// TIA Portal V20 export
DATA_BLOCK "DB_Stoermeldungen"   // DB512
TITLE = Schnittstelle OP_AG 1
{ S7_Optimized_Access := 'FALSE' }
AUTHOR : SD
FAMILY : KOMM
// stored: AutoNumber false
   VAR RETAIN
      Allgemeine { S7_SetPoint := 'True'} : "Störmeldung";
      Allgemeine_1 { S7_SetPoint := 'True'} : "Störmeldung";
      SM_Wartungszähler { S7_SetPoint := 'True'} : "Störmeldung";
      Störmeldungen_PN : "Störmeldung_PN";
   END_VAR
BEGIN
   Allgemeine.Störmeldung[0] := FALSE;
   Allgemeine.Störmeldung[1] := FALSE;   // SM1 Systemdruck nicht vorhanden ! Prüfen und Weiter mit ACK
   Allgemeine.Störmeldung[2] := FALSE;   // SM2 Anlagendruck nicht aufgebaut -939S1
   Allgemeine.Störmeldung[3] := FALSE;   // SM3 Algemein Richten Gesamtanlage erforderlich
   Allgemeine.Störmeldung[4] := FALSE;   // SM4 Richten Gesamtanlage nach Teil neu geladen
   Allgemeine.Störmeldung[5] := FALSE;   // SM5
   Allgemeine.Störmeldung[6] := FALSE;   // SM6
   Allgemeine.Störmeldung[7] := FALSE;   // SM7
   Allgemeine.Störmeldung[8] := FALSE;   // SM8
   Allgemeine.Störmeldung[9] := FALSE;   // SM9
   Allgemeine.Störmeldung[10] := FALSE;   // SM10
   Allgemeine.Störmeldung[11] := FALSE;   // SM11
   Allgemeine.Störmeldung[12] := FALSE;   // SM12
   Allgemeine.Störmeldung[13] := FALSE;   // SM13
   Allgemeine.Störmeldung[14] := FALSE;   // SM14
   Allgemeine.Störmeldung[15] := FALSE;   // SM15
   Allgemeine.Störmeldung[16] := FALSE;   // SM16
   Allgemeine.Störmeldung[17] := FALSE;   // SM17
   Allgemeine.Störmeldung[18] := FALSE;   // SM18
   Allgemeine.Störmeldung[19] := FALSE;   // SM19
   Allgemeine.Störmeldung[20] := FALSE;   // SM20
   Allgemeine.Störmeldung[21] := FALSE;   // SM21
   Allgemeine.Störmeldung[22] := FALSE;   // SM22
   Allgemeine.Störmeldung[23] := FALSE;   // SM23
   Allgemeine.Störmeldung[24] := FALSE;   // SM24
   Allgemeine.Störmeldung[25] := FALSE;   // SM25
   Allgemeine.Störmeldung[26] := FALSE;   // SM26
   Allgemeine.Störmeldung[27] := FALSE;   // SM27
   Allgemeine.Störmeldung[28] := FALSE;   // SM28
   Allgemeine.Störmeldung[29] := FALSE;   // SM29
   Allgemeine.Störmeldung[30] := FALSE;   // SM30
   Allgemeine.Störmeldung[31] := FALSE;   // SM31
   Allgemeine_1.Störmeldung[0] := FALSE;   // SM32 Schutztüre 1 nicht verriegelt
   Allgemeine_1.Störmeldung[1] := FALSE;   // SM33 Schutztüre 2 nicht verriegelt
   Allgemeine_1.Störmeldung[2] := FALSE;   // SM34 Schutztüre 3 nicht verriegelt
   Allgemeine_1.Störmeldung[3] := FALSE;   // SM35 Schutztüre 4 nicht verriegelt
   Allgemeine_1.Störmeldung[4] := FALSE;   // SM36 Schutztüre 5 nicht verriegelt
   Allgemeine_1.Störmeldung[5] := FALSE;   // SM37 Schutztüre 6 nicht verriegelt
   Allgemeine_1.Störmeldung[6] := FALSE;   // SM38 Schutztüre 7 nicht verriegelt
   Allgemeine_1.Störmeldung[7] := FALSE;   // SM39 Schutztüre 8 nicht verriegelt
   Allgemeine_1.Störmeldung[8] := FALSE;   // SM40 Schutztüre 9 nicht verriegelt
   Allgemeine_1.Störmeldung[9] := FALSE;   // SM41 Schutztüre 10 nicht verriegelt
   Allgemeine_1.Störmeldung[10] := FALSE;   // SM42 Schutztüre 11 nicht verriegelt
   Allgemeine_1.Störmeldung[11] := FALSE;   // SM43 Steuerspannung 24V nicht in Ordnung
   Allgemeine_1.Störmeldung[12] := FALSE;   // SM44 Not-Aus Taster Bedienpanel
   Allgemeine_1.Störmeldung[13] := FALSE;   // SM45 Not-Aus Taster extern
   Allgemeine_1.Störmeldung[14] := FALSE;   // SM46 Kontrolle Box 1 voll -> leeren -> Start
   Allgemeine_1.Störmeldung[15] := FALSE;   // SM47 Kontrolle Box 2 voll -> leeren -> Start
   Allgemeine_1.Störmeldung[16] := FALSE;   // SM48 Kontrolle Box 3 voll -> leeren -> Start
   Allgemeine_1.Störmeldung[17] := FALSE;   // SM49 NIO Box 1 voll -> leeren -> Start
   Allgemeine_1.Störmeldung[18] := FALSE;   // SM50 NIO Box 2 voll -> leeren -> Start
   Allgemeine_1.Störmeldung[19] := FALSE;   // SM51 IO Box voll -> leeren -> Start
   Allgemeine_1.Störmeldung[20] := FALSE;   // SM52 Teiledaten wurden nicht richtig übertragen
   Allgemeine_1.Störmeldung[21] := FALSE;   // SM53 IO Box in Einhausung voll -> leeren -> Start
   Allgemeine_1.Störmeldung[22] := FALSE;   // SM54
   Allgemeine_1.Störmeldung[23] := FALSE;   // SM55 Anlagendruck bei Not-Halt nicht abgebaut -939S2
   Allgemeine_1.Störmeldung[24] := FALSE;   // SM56 Überspannungsschutz nicht OK
   Allgemeine_1.Störmeldung[25] := FALSE;   // SM57
   Allgemeine_1.Störmeldung[26] := FALSE;   // SM58
   Allgemeine_1.Störmeldung[27] := FALSE;   // SM59
   Allgemeine_1.Störmeldung[28] := FALSE;   // SM60
   Allgemeine_1.Störmeldung[29] := FALSE;   // SM61
   Allgemeine_1.Störmeldung[30] := FALSE;   // SM62
   Allgemeine_1.Störmeldung[31] := FALSE;   // SM63
   SM_Wartungszähler.Störmeldung[0] := FALSE;   // SM576 Wartungszähler 1
   SM_Wartungszähler.Störmeldung[1] := FALSE;   // SM577 Wartungszähler 2
   SM_Wartungszähler.Störmeldung[2] := FALSE;   // SM578 Wartungszähler 3
   SM_Wartungszähler.Störmeldung[3] := FALSE;   // SM579 Wartungszähler 4
   SM_Wartungszähler.Störmeldung[4] := FALSE;   // SM580 Wartungszähler 5
   SM_Wartungszähler.Störmeldung[5] := FALSE;   // SM581 Wartungszähler 6
   SM_Wartungszähler.Störmeldung[6] := FALSE;   // SM582 Wartungszähler 7
   SM_Wartungszähler.Störmeldung[7] := FALSE;   // SM583
   SM_Wartungszähler.Störmeldung[8] := FALSE;   // SM584
   SM_Wartungszähler.Störmeldung[9] := FALSE;   // SM585
   SM_Wartungszähler.Störmeldung[10] := FALSE;   // SM586
   SM_Wartungszähler.Störmeldung[11] := FALSE;   // SM587
   SM_Wartungszähler.Störmeldung[12] := FALSE;   // SM588
   SM_Wartungszähler.Störmeldung[13] := FALSE;   // SM589
   SM_Wartungszähler.Störmeldung[14] := FALSE;   // SM590
   SM_Wartungszähler.Störmeldung[15] := FALSE;   // SM591
   SM_Wartungszähler.Störmeldung[16] := FALSE;   // SM592
   SM_Wartungszähler.Störmeldung[17] := FALSE;   // SM593
   SM_Wartungszähler.Störmeldung[18] := FALSE;   // SM594
   SM_Wartungszähler.Störmeldung[19] := FALSE;   // SM595
   SM_Wartungszähler.Störmeldung[20] := FALSE;   // SM596
   SM_Wartungszähler.Störmeldung[21] := FALSE;   // SM597
   SM_Wartungszähler.Störmeldung[22] := FALSE;   // SM598
   SM_Wartungszähler.Störmeldung[23] := FALSE;   // SM599
   SM_Wartungszähler.Störmeldung[24] := FALSE;   // SM600
   SM_Wartungszähler.Störmeldung[25] := FALSE;   // SM601
   SM_Wartungszähler.Störmeldung[26] := FALSE;   // SM602
   SM_Wartungszähler.Störmeldung[27] := FALSE;   // SM603
   SM_Wartungszähler.Störmeldung[28] := FALSE;   // SM604
   SM_Wartungszähler.Störmeldung[29] := FALSE;   // SM605
   SM_Wartungszähler.Störmeldung[30] := FALSE;   // SM606
   SM_Wartungszähler.Störmeldung[31] := FALSE;   // SM607
   Störmeldungen_PN.Störmeldung_PN[0] := FALSE;   // SM608 Sammelstörung Profinet
   Störmeldungen_PN.Störmeldung_PN[1] := FALSE;   // SM609 Ausfall/Störung +HS1-101A1 Pluto Gateway Profinet
   Störmeldungen_PN.Störmeldung_PN[2] := FALSE;   // SM610 Ausfall/Störung +HS1-41T1 Pos 3.0 Drehteller
   Störmeldungen_PN.Störmeldung_PN[3] := FALSE;   // SM611 Ausfall/Störung +HS1-43T1 Pos 3.1 Rutsche Anschlag Oriental E-Antrieb
   Störmeldungen_PN.Störmeldung_PN[4] := FALSE;   // SM612 Ausfall/Störung +HS1-44T1 Pos 3.1 Spannvorrichtung LinMot
   Störmeldungen_PN.Störmeldung_PN[5] := FALSE;   // SM613 Ausfall/Störung +HS1-46T1 Pos 3.3 Ausdrehen Oriental E-Antrieb
   Störmeldungen_PN.Störmeldung_PN[6] := FALSE;   // SM614 Ausfall/Störung +HS1-50T1 Pos 3.7 Ausdrehen Oriental E-Antrieb
   Störmeldungen_PN.Störmeldung_PN[7] := FALSE;   // SM615 Ausfall/Störung +HS1-55T1 Pos 3.11 Spannvorrichtung LinMot
   Störmeldungen_PN.Störmeldung_PN[8] := FALSE;   // SM616 Ausfall/Störung +Feld-941ZX1-943ZX1 Multipolverteiler 1-3
   Störmeldungen_PN.Störmeldung_PN[9] := FALSE;   // SM617 Ausfall/Störung +Feld-961VB1 Ventilblock 1
   Störmeldungen_PN.Störmeldung_PN[10] := FALSE;   // SM618 Ausfall/Störung -1131A1 POS 3.1 Epson Roboter
   Störmeldungen_PN.Störmeldung_PN[11] := FALSE;   // SM619 Ausfall/Störung -2131A1 POS 3.11 Epson Roboter
   Störmeldungen_PN.Störmeldung_PN[12] := FALSE;   // SM620 Ausfall/Störung
   Störmeldungen_PN.Störmeldung_PN[13] := FALSE;   // SM621 Ausfall/Störung
   Störmeldungen_PN.Störmeldung_PN[14] := FALSE;   // SM622 Ausfall/Störung
   Störmeldungen_PN.Störmeldung_PN[15] := FALSE;   // SM623 Ausfall/Störung
   Störmeldungen_PN.Störmeldung_PN[16] := FALSE;   // SM624 Ausfall/Störung
   Störmeldungen_PN.Störmeldung_PN[17] := FALSE;   // SM625 Ausfall/Störung
   Störmeldungen_PN.Störmeldung_PN[18] := FALSE;   // SM626 Ausfall/Störung
   Störmeldungen_PN.Störmeldung_PN[19] := FALSE;   // SM627 Ausfall/Störung
   Störmeldungen_PN.Störmeldung_PN[20] := FALSE;   // SM628 Ausfall/Störung
   Störmeldungen_PN.Störmeldung_PN[21] := FALSE;   // SM629 Ausfall/Störung
   Störmeldungen_PN.Störmeldung_PN[22] := FALSE;   // SM630 Ausfall/Störung
   Störmeldungen_PN.Störmeldung_PN[23] := FALSE;   // SM631 Ausfall/Störung
   Störmeldungen_PN.Störmeldung_PN[24] := FALSE;   // SM632 Ausfall/Störung
   Störmeldungen_PN.Störmeldung_PN[25] := FALSE;   // SM633 Ausfall/Störung
   Störmeldungen_PN.Störmeldung_PN[26] := FALSE;   // SM634 Ausfall/Störung
   Störmeldungen_PN.Störmeldung_PN[27] := FALSE;   // SM635 Ausfall/Störung
   Störmeldungen_PN.Störmeldung_PN[28] := FALSE;   // SM636 Ausfall/Störung
   Störmeldungen_PN.Störmeldung_PN[29] := FALSE;   // SM637 Ausfall/Störung
   Störmeldungen_PN.Störmeldung_PN[30] := FALSE;   // SM638 Ausfall/Störung
   Störmeldungen_PN.Störmeldung_PN[31] := FALSE;   // SM639 Ausfall/Störung
   Störmeldungen_PN.Störmeldung_PN[32] := FALSE;   // SM640 Ausfall/Störung
   Störmeldungen_PN.Störmeldung_PN[33] := FALSE;   // SM641 Ausfall/Störung
   Störmeldungen_PN.Störmeldung_PN[34] := FALSE;   // SM642 Ausfall/Störung
   Störmeldungen_PN.Störmeldung_PN[35] := FALSE;   // SM643 Ausfall/Störung
   Störmeldungen_PN.Störmeldung_PN[36] := FALSE;   // SM644 Ausfall/Störung
   Störmeldungen_PN.Störmeldung_PN[37] := FALSE;   // SM645 Ausfall/Störung
   Störmeldungen_PN.Störmeldung_PN[38] := FALSE;   // SM646 Ausfall/Störung
   Störmeldungen_PN.Störmeldung_PN[39] := FALSE;   // SM647 Ausfall/Störung
   Störmeldungen_PN.Störmeldung_PN[40..127] := FALSE;
END_DATA_BLOCK
